// TIA Portal V17 export
FUNCTION "FC_T04a_TON_DB" : Void   // FC141, LAD
{ S7_Optimized_Access := 'TRUE' }
// stored: SetENOAutomatically false
   VAR_INPUT
      Demarrer : Bool;
   END_VAR
   VAR_OUTPUT
      Tempo_OK : Bool;
   END_VAR
BEGIN

REGION Network 1: TON avec DB d'instance
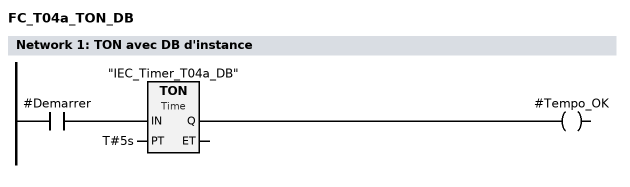
   RUNG wire#powerrail
      Contact( #Demarrer )
      { S7_Templates := "time_type := Time" } "IEC_Timer_T04a_DB".TON(pt := T#5s, et =>)
      Coil( #Tempo_OK )
   END_RUNG
   // the same network as SCL:
   "IEC_Timer_T04a_DB".TON(IN := #Demarrer, PT := T#5s);
   #Tempo_OK := "IEC_Timer_T04a_DB".Q;
END_REGION
END_FUNCTION
